Yaskawa INFORM job: MANPRO_REV_2.JBI

/JOB
//NAME MANPRO_REV_2
//POS
///NPOS 15,0,15,0,0,0
///TOOL 0
///POSTYPE PULSE
///PULSE
C00000=-729,-59979,-60060,-74,-89734,186
C00001=3819,16382,-27236,870,-54500,42809
C00002=3525,16854,-28349,958,-53276,42967
C00003=-3358,28738,-45607,-1245,-29542,40340
C00004=-8926,39935,-26267,5691,-33626,4077
C00005=-16606,45376,-17783,5613,-43931,-15629
C00006=-16077,39808,-21056,7196,-36422,-13209
C00007=-21057,8484,-56828,1119,-11848,1649
C00008=-22681,18094,-67654,2450,7059,-6589
C00009=-16365,16976,-69325,-17660,7079,1120
C00010=-17296,-5027,-68711,-157,-1378,-2962
C00011=-21413,17494,-103035,-1830,53788,-17035
C00012=-19881,21209,-97135,-2963,52531,-16955
C00013=-4537,-41986,-65927,19082,-22840,-20309
C00014=-1,-60103,-60032,2,-90053,2
EC00000=1
EC00001=-82435
EC00002=-69446
EC00003=-1216
EC00004=-1216
EC00005=-1216
EC00006=-22347
EC00007=-82435
EC00008=-82435
EC00009=-82435
EC00010=-82435
EC00011=-160520
EC00012=-160520
EC00013=-80844
EC00014=-1644
//INST
///DATE 2026/04/27 12:40
///ATTR SC,RW
///GROUP1 RB1,ST1
NOP
MOVL C00000 EC00000 V=833.3
MOVL C00001 EC00001 V=833.3
MOVL C00002 EC00002 V=83.3
MOVC C00003 EC00003 V=83.3
ARCON ASF#(2)
MOVC C00004 EC00004 V=4.7
MOVC C00005 EC00005 V=5.0
ARCOF AEF#(2)
MOVL C00006 EC00006 V=83.3
MOVL C00007 EC00007 V=83.3
MOVL C00008 EC00008 V=83.3
ARCON ASF#(2)
MOVL C00009 EC00009 V=3.3
ARCOF AEF#(2)
MOVL C00010 EC00010 V=333.3
MOVL C00011 EC00011 V=50.0
ARCON ASF#(2)
MOVL C00012 EC00012 V=4.8
ARCOF AEF#(2)
MOVL C00013 EC00013 V=333.3
MOVL C00014 EC00014 V=333.3
CALL JOB:CLEAN_R1
END
